{attribute 'qualified_only'}
{attribute 'strict'}
{attribute 'to_string'}
TYPE E_PackMLStates :
(
	Idle := 0,
	Starting, 
	Execute, 
	Suspending, 
	Suspended, 
	Unsuspending, 
	Holding,
	Held,
	Unholding,
	Resetting,
	Aborting,
	Aborted, 
	Clearing,
	Stopping,
	Stopped
);
END_TYPE

(* stored: Version 1.1.0.1
   DUT E_PackMLStates: Id {8662dd63-e7b9-4231-9ff0-533ef6ce4f51} *)
